// TIA Portal V20 export
TYPE "TDiag_StatusExt"
   STRUCT
      Interfaceld : HW_ANY;
      ID : CONN_OUC;
      ConnectionType : Byte;
      ActivateEstablished : Bool;
      State : Byte;
      Kind : Byte;
      SentBytes : UDInt;
      ReceivedBytes : UDInt;
   END_STRUCT;
END_TYPE
